(* IEC 61131-3 sources: trust-platform/examples/OSCAT/district_pump_network_proxy_mediator/oop/src, 3 files *)

(* ---- Main.st ---- *)
(* Pattern role: IStationProxy is the contract boundary for the Proxy and Mediator example. *)
INTERFACE IStationProxy
    PROPERTY StationId : INT
    GET
    END_GET
    END_PROPERTY

    PROPERTY DemandM3H : REAL
    GET
    END_GET
    END_PROPERTY

    PROPERTY IsStale : BOOL
    GET
    END_GET
    END_PROPERTY

    PROPERTY QualityGood : BOOL
    GET
    END_GET
    END_PROPERTY

    METHOD UpdateProxy
    VAR_INPUT
        DemandM3H : REAL;
        QualityGoodInput : BOOL;
        AgeSeconds : INT;
    END_VAR
    END_METHOD
END_INTERFACE

(* Pattern role: LocalStationProxy is a concrete implementation in the Proxy and Mediator example. *)
FUNCTION_BLOCK LocalStationProxy IMPLEMENTS IStationProxy
VAR
    DemandValue : REAL;
END_VAR

METHOD PUBLIC UpdateProxy
VAR_INPUT
    DemandM3H : REAL;
    QualityGoodInput : BOOL;
    AgeSeconds : INT;
END_VAR
DemandValue := DemandM3H;
END_METHOD

PUBLIC PROPERTY StationId : INT
GET
    StationId := INT#0;
END_GET
END_PROPERTY

PUBLIC PROPERTY DemandM3H : REAL
GET
    DemandM3H := DemandValue;
END_GET
END_PROPERTY

PUBLIC PROPERTY IsStale : BOOL
GET
    IsStale := FALSE;
END_GET
END_PROPERTY

PUBLIC PROPERTY QualityGood : BOOL
GET
    QualityGood := TRUE;
END_GET
END_PROPERTY
END_FUNCTION_BLOCK

(* Pattern role: RemoteStationProxy is a concrete implementation in the Proxy and Mediator example. *)
FUNCTION_BLOCK RemoteStationProxy IMPLEMENTS IStationProxy
VAR
    StationIdValue : INT;
    DemandValue : REAL;
    StaleValue : BOOL;
    QualityGoodValue : BOOL;
    LastAgeSecondsValue : INT;
END_VAR

METHOD PUBLIC Configure
VAR_INPUT
    StationId : INT;
END_VAR
StationIdValue := StationId;
END_METHOD

METHOD PUBLIC UpdateProxy
VAR_INPUT
    DemandM3H : REAL;
    QualityGoodInput : BOOL;
    AgeSeconds : INT;
END_VAR
DemandValue := DemandM3H;
QualityGoodValue := QualityGoodInput;
LastAgeSecondsValue := AgeSeconds;
StaleValue := (NOT QualityGoodInput) OR (AgeSeconds > INT#30);
END_METHOD

PUBLIC PROPERTY StationId : INT
GET
    StationId := StationIdValue;
END_GET
END_PROPERTY

PUBLIC PROPERTY DemandM3H : REAL
GET
    DemandM3H := DemandValue;
END_GET
END_PROPERTY

PUBLIC PROPERTY IsStale : BOOL
GET
    IsStale := StaleValue;
END_GET
END_PROPERTY

PUBLIC PROPERTY QualityGood : BOOL
GET
    QualityGood := QualityGoodValue;
END_GET
END_PROPERTY

PUBLIC PROPERTY LastAgeSeconds : INT
GET
    LastAgeSeconds := LastAgeSecondsValue;
END_GET
END_PROPERTY
END_FUNCTION_BLOCK

(* Composition role: DemandMediator owns the collaborating objects used by this Proxy and Mediator example. *)
FUNCTION_BLOCK DemandMediator
VAR
    Local : LocalStationProxy;
    NorthRemote : RemoteStationProxy;
    EastRemote : RemoteStationProxy;
    TotalDemandM3HValue : REAL;
    PumpSpeedPctValue : REAL;
    RemoteStaleCountValue : INT;
    ClassAAlarmValue : BOOL;
END_VAR

METHOD PUBLIC Initialize
NorthRemote.Configure(StationId := INT#1);
EastRemote.Configure(StationId := INT#2);
END_METHOD

METHOD PRIVATE AcceptProxy
VAR_INPUT
    Station : IStationProxy;
    CountStale : BOOL;
END_VAR
IF Station.IsStale THEN
    IF CountStale THEN
        RemoteStaleCountValue := RemoteStaleCountValue + INT#1;
    END_IF;
ELSE
    TotalDemandM3HValue := TotalDemandM3HValue + Station.DemandM3H;
END_IF;
END_METHOD

METHOD PUBLIC Update : REAL
VAR_INPUT
    LocalDemandM3H : REAL;
    NorthDemandM3H : REAL;
    NorthQualityGood : BOOL;
    NorthAgeSeconds : INT;
    EastDemandM3H : REAL;
    EastQualityGood : BOOL;
    EastAgeSeconds : INT;
    SuctionHealthy : BOOL;
END_VAR
Local.UpdateProxy(DemandM3H := LocalDemandM3H, QualityGoodInput := TRUE, AgeSeconds := INT#0);
NorthRemote.UpdateProxy(DemandM3H := NorthDemandM3H, QualityGoodInput := NorthQualityGood, AgeSeconds := NorthAgeSeconds);
EastRemote.UpdateProxy(DemandM3H := EastDemandM3H, QualityGoodInput := EastQualityGood, AgeSeconds := EastAgeSeconds);

TotalDemandM3HValue := REAL#0.0;
RemoteStaleCountValue := INT#0;
AcceptProxy(Station := Local, CountStale := FALSE);
AcceptProxy(Station := NorthRemote, CountStale := TRUE);
AcceptProxy(Station := EastRemote, CountStale := TRUE);

ClassAAlarmValue := NOT SuctionHealthy;
IF ClassAAlarmValue THEN
    PumpSpeedPctValue := REAL#0.0;
ELSE
    PumpSpeedPctValue := LIMIT(REAL#0.0, TotalDemandM3HValue * REAL#2.0, REAL#100.0);
END_IF;
Update := PumpSpeedPctValue;
END_METHOD

PUBLIC PROPERTY TotalDemandM3H : REAL
GET
    TotalDemandM3H := TotalDemandM3HValue;
END_GET
END_PROPERTY

PUBLIC PROPERTY PumpSpeedPct : REAL
GET
    PumpSpeedPct := PumpSpeedPctValue;
END_GET
END_PROPERTY

PUBLIC PROPERTY RemoteStaleCount : INT
GET
    RemoteStaleCount := RemoteStaleCountValue;
END_GET
END_PROPERTY

PUBLIC PROPERTY ClassAAlarm : BOOL
GET
    ClassAAlarm := ClassAAlarmValue;
END_GET
END_PROPERTY
END_FUNCTION_BLOCK

(* Scan role: Main wires the example objects and exposes the PLC call path under test. *)
PROGRAM Main
VAR
    Network : DemandMediator;
    LocalDemandRaw : INT;
    NorthDemandRaw : INT;
    EastDemandRaw : INT;
    NorthAgeSeconds : INT;
    EastAgeSeconds : INT;
    NorthQualityGood : BOOL;
    EastQualityGood : BOOL;
    SuctionHealthy : BOOL;
    PumpSpeedRaw : INT;
    StaleAlarmOut : BOOL;
END_VAR
Network.Initialize();
Network.Update(LocalDemandM3H := INT_TO_REAL(LocalDemandRaw), NorthDemandM3H := INT_TO_REAL(NorthDemandRaw), NorthQualityGood := NorthQualityGood, NorthAgeSeconds := NorthAgeSeconds, EastDemandM3H := INT_TO_REAL(EastDemandRaw), EastQualityGood := EastQualityGood, EastAgeSeconds := EastAgeSeconds, SuctionHealthy := SuctionHealthy);
PumpSpeedRaw := REAL_TO_INT(Network.PumpSpeedPct);
StaleAlarmOut := Network.RemoteStaleCount > INT#0;
END_PROGRAM

(* ---- Configuration.st ---- *)
CONFIGURATION DistrictPumpNetworkProxyMediatorOopConfiguration
RESOURCE DistrictPumpNetworkProxyMediatorOop ON PLC
    TASK MainTask (INTERVAL := T#100ms, PRIORITY := 1);
    PROGRAM Network WITH MainTask : Main;
END_RESOURCE
VAR_CONFIG
    Network.LocalDemandRaw AT %IW2 : INT;
    Network.NorthDemandRaw AT %IW4 : INT;
    Network.EastDemandRaw AT %IW6 : INT;
    Network.NorthAgeSeconds AT %IW8 : INT;
    Network.EastAgeSeconds AT %IW10 : INT;
    Network.NorthQualityGood AT %IX0.0 : BOOL;
    Network.EastQualityGood AT %IX0.1 : BOOL;
    Network.SuctionHealthy AT %IX0.2 : BOOL;
    Network.PumpSpeedRaw AT %QW2 : INT;
    Network.StaleAlarmOut AT %QX0.0 : BOOL;
END_VAR
END_CONFIGURATION

(* ---- Tests.st ---- *)
TEST_PROGRAM DistrictMediatorBalancesHealthyRemoteDemand
VAR
    Network : DemandMediator;
END_VAR

Network.Initialize();
ASSERT_EQUAL(EXPECTED := REAL#90.0, ACTUAL := Network.Update(LocalDemandM3H := REAL#20.0, NorthDemandM3H := REAL#15.0, NorthQualityGood := TRUE, NorthAgeSeconds := INT#5, EastDemandM3H := REAL#10.0, EastQualityGood := TRUE, EastAgeSeconds := INT#5, SuctionHealthy := TRUE));
ASSERT_EQUAL(EXPECTED := REAL#45.0, ACTUAL := Network.TotalDemandM3H);
ASSERT_EQUAL(EXPECTED := INT#0, ACTUAL := Network.RemoteStaleCount);
END_TEST_PROGRAM

TEST_PROGRAM DistrictProxyDropsStaleRemoteDemand
VAR
    Network : DemandMediator;
END_VAR

Network.Initialize();
ASSERT_EQUAL(EXPECTED := REAL#40.0, ACTUAL := Network.Update(LocalDemandM3H := REAL#20.0, NorthDemandM3H := REAL#15.0, NorthQualityGood := TRUE, NorthAgeSeconds := INT#45, EastDemandM3H := REAL#10.0, EastQualityGood := FALSE, EastAgeSeconds := INT#5, SuctionHealthy := TRUE));
ASSERT_EQUAL(EXPECTED := REAL#20.0, ACTUAL := Network.TotalDemandM3H);
ASSERT_EQUAL(EXPECTED := INT#2, ACTUAL := Network.RemoteStaleCount);
END_TEST_PROGRAM

TEST_PROGRAM DistrictMediatorTripsOnLocalSuctionLoss
VAR
    Network : DemandMediator;
END_VAR

Network.Initialize();
ASSERT_EQUAL(EXPECTED := REAL#0.0, ACTUAL := Network.Update(LocalDemandM3H := REAL#20.0, NorthDemandM3H := REAL#15.0, NorthQualityGood := TRUE, NorthAgeSeconds := INT#5, EastDemandM3H := REAL#10.0, EastQualityGood := TRUE, EastAgeSeconds := INT#5, SuctionHealthy := FALSE));
ASSERT_TRUE(IN := Network.ClassAAlarm);
END_TEST_PROGRAM

(* Multi-scan proxy-aging test: drives the same network through
   healthy, stale, and recovered remote states. Catches bugs where
   RemoteStaleCount stays sticky after recovery, or where a stale
   remote's last-known demand keeps contributing to TotalDemandM3H. *)
TEST_PROGRAM DistrictProxyTracksFreshAndStaleStateAcrossScans
VAR
    Network : DemandMediator;
END_VAR

Network.Initialize();

(* Scan 1: both remotes fresh *)
Network.Update(LocalDemandM3H := REAL#20.0, NorthDemandM3H := REAL#15.0, NorthQualityGood := TRUE, NorthAgeSeconds := INT#5, EastDemandM3H := REAL#10.0, EastQualityGood := TRUE, EastAgeSeconds := INT#5, SuctionHealthy := TRUE);
ASSERT_EQUAL(EXPECTED := INT#0, ACTUAL := Network.RemoteStaleCount);

(* Scan 2: north stale, east bad-quality *)
Network.Update(LocalDemandM3H := REAL#20.0, NorthDemandM3H := REAL#15.0, NorthQualityGood := TRUE, NorthAgeSeconds := INT#45, EastDemandM3H := REAL#10.0, EastQualityGood := FALSE, EastAgeSeconds := INT#5, SuctionHealthy := TRUE);
ASSERT_EQUAL(EXPECTED := INT#2, ACTUAL := Network.RemoteStaleCount);

(* Scan 3: both remotes recover - stale count must reset to zero *)
Network.Update(LocalDemandM3H := REAL#20.0, NorthDemandM3H := REAL#15.0, NorthQualityGood := TRUE, NorthAgeSeconds := INT#5, EastDemandM3H := REAL#10.0, EastQualityGood := TRUE, EastAgeSeconds := INT#5, SuctionHealthy := TRUE);
ASSERT_EQUAL(EXPECTED := INT#0, ACTUAL := Network.RemoteStaleCount);
ASSERT_EQUAL(EXPECTED := REAL#45.0, ACTUAL := Network.TotalDemandM3H);
END_TEST_PROGRAM

(* Boundary: exact age threshold. The proxy uses AgeSeconds > 30 as
   the staleness rule, so 30 is fresh, 31 is stale. *)
TEST_PROGRAM DistrictProxyAgeBoundaryAtExactThirty
VAR
    Network : DemandMediator;
END_VAR

Network.Initialize();

(* Age = 30 (exact threshold, still fresh by > rule) *)
Network.Update(LocalDemandM3H := REAL#10.0, NorthDemandM3H := REAL#5.0, NorthQualityGood := TRUE, NorthAgeSeconds := INT#30, EastDemandM3H := REAL#0.0, EastQualityGood := TRUE, EastAgeSeconds := INT#0, SuctionHealthy := TRUE);
ASSERT_EQUAL(EXPECTED := INT#0, ACTUAL := Network.RemoteStaleCount);
ASSERT_EQUAL(EXPECTED := REAL#15.0, ACTUAL := Network.TotalDemandM3H);

(* Age = 31 (over threshold, stale) *)
Network.Update(LocalDemandM3H := REAL#10.0, NorthDemandM3H := REAL#5.0, NorthQualityGood := TRUE, NorthAgeSeconds := INT#31, EastDemandM3H := REAL#0.0, EastQualityGood := TRUE, EastAgeSeconds := INT#0, SuctionHealthy := TRUE);
ASSERT_EQUAL(EXPECTED := INT#1, ACTUAL := Network.RemoteStaleCount);
ASSERT_EQUAL(EXPECTED := REAL#10.0, ACTUAL := Network.TotalDemandM3H);
END_TEST_PROGRAM

(* RemoteStationProxy in isolation: tests the staleness rule
   directly on a single proxy, verifies the IsStale property tracks
   the rule (NOT QualityGood OR AgeSeconds > 30). *)
TEST_PROGRAM DistrictRemoteProxyStalenessRuleInIsolation
VAR
    Remote : RemoteStationProxy;
END_VAR

Remote.Configure(StationId := INT#42);
ASSERT_EQUAL(EXPECTED := INT#42, ACTUAL := Remote.StationId);

(* Healthy: fresh demand, good quality *)
Remote.UpdateProxy(DemandM3H := REAL#7.5, QualityGoodInput := TRUE, AgeSeconds := INT#10);
ASSERT_FALSE(IN := Remote.IsStale);
ASSERT_TRUE(IN := Remote.QualityGood);
ASSERT_NEAR(EXPECTED := REAL#7.5, ACTUAL := Remote.DemandM3H, DELTA := REAL#0.001);

(* Aged out *)
Remote.UpdateProxy(DemandM3H := REAL#7.5, QualityGoodInput := TRUE, AgeSeconds := INT#100);
ASSERT_TRUE(IN := Remote.IsStale);

(* Bad quality even at age 0 *)
Remote.UpdateProxy(DemandM3H := REAL#7.5, QualityGoodInput := FALSE, AgeSeconds := INT#0);
ASSERT_TRUE(IN := Remote.IsStale);

(* Recovered *)
Remote.UpdateProxy(DemandM3H := REAL#5.0, QualityGoodInput := TRUE, AgeSeconds := INT#5);
ASSERT_FALSE(IN := Remote.IsStale);
END_TEST_PROGRAM

(* LocalStationProxy is never stale by design - the local PLC's own
   scan tags do not have a freshness contract. *)
TEST_PROGRAM DistrictLocalProxyIsNeverStale
VAR
    Local : LocalStationProxy;
END_VAR

(* Exercising UpdateProxy with bad quality and stale age must not flip IsStale *)
Local.UpdateProxy(DemandM3H := REAL#42.0, QualityGoodInput := FALSE, AgeSeconds := INT#9999);
ASSERT_FALSE(IN := Local.IsStale);
ASSERT_TRUE(IN := Local.QualityGood);
ASSERT_EQUAL(EXPECTED := INT#0, ACTUAL := Local.StationId);
ASSERT_NEAR(EXPECTED := REAL#42.0, ACTUAL := Local.DemandM3H, DELTA := REAL#0.001);
END_TEST_PROGRAM

(* Suction trip overrides aggregated demand: even with all stations
   healthy, ClassA alarm forces PumpSpeed = 0. *)
TEST_PROGRAM DistrictSuctionTripOverridesHealthyAggregate
VAR
    Network : DemandMediator;
END_VAR

Network.Initialize();

(* All healthy except suction *)
ASSERT_EQUAL(EXPECTED := REAL#0.0, ACTUAL := Network.Update(LocalDemandM3H := REAL#20.0, NorthDemandM3H := REAL#15.0, NorthQualityGood := TRUE, NorthAgeSeconds := INT#5, EastDemandM3H := REAL#10.0, EastQualityGood := TRUE, EastAgeSeconds := INT#5, SuctionHealthy := FALSE));
ASSERT_TRUE(IN := Network.ClassAAlarm);
(* TotalDemand should still aggregate (mediator computes both) *)
ASSERT_EQUAL(EXPECTED := REAL#45.0, ACTUAL := Network.TotalDemandM3H);

(* Recovery: suction comes back, command resumes *)
ASSERT_EQUAL(EXPECTED := REAL#90.0, ACTUAL := Network.Update(LocalDemandM3H := REAL#20.0, NorthDemandM3H := REAL#15.0, NorthQualityGood := TRUE, NorthAgeSeconds := INT#5, EastDemandM3H := REAL#10.0, EastQualityGood := TRUE, EastAgeSeconds := INT#5, SuctionHealthy := TRUE));
ASSERT_FALSE(IN := Network.ClassAAlarm);
END_TEST_PROGRAM

(* Pump speed clamps at 100% even with very large total demand. *)
TEST_PROGRAM DistrictPumpSpeedSaturatesAtHundredPercent
VAR
    Network : DemandMediator;
END_VAR

Network.Initialize();

(* Total demand 200 m3/h * 2 = 400; clamped to 100 *)
ASSERT_EQUAL(EXPECTED := REAL#100.0, ACTUAL := Network.Update(LocalDemandM3H := REAL#100.0, NorthDemandM3H := REAL#50.0, NorthQualityGood := TRUE, NorthAgeSeconds := INT#5, EastDemandM3H := REAL#50.0, EastQualityGood := TRUE, EastAgeSeconds := INT#5, SuctionHealthy := TRUE));
ASSERT_EQUAL(EXPECTED := REAL#200.0, ACTUAL := Network.TotalDemandM3H);
END_TEST_PROGRAM
